{attribute 'qualified_only'}
VAR_GLOBAL
	//Inputs
	DI_E0_0     AT%I*	:BOOL;
	DI_E0_1		AT%I*	:BOOL;
	
	DI_E50_0	AT%I*	:BOOL;
	DI_E50_1	AT%I*	:BOOL;
	DI_E50_2	AT%I*	:BOOL;
	
	DI_E1050_0	AT%I*	:BOOL;
	DI_E1050_1	AT%I*	:BOOL;
	DI_E1050_2	AT%I*	:BOOL;
	DI_E1050_3	AT%I*	:BOOL;
	DI_E1050_4	AT%I*	:BOOL;
	DI_E1050_5	AT%I*	:BOOL;
	
	DI_E1051_0	AT%I*	:BOOL;
	DI_E1051_1	AT%I*	:BOOL;
	DI_E1051_2	AT%I*	:BOOL;
	DI_E1051_3	AT%I*	:BOOL;
	
	DI_E1052_0	AT%I*	:BOOL;
	DI_E1052_1	AT%I*	:BOOL;
	DI_E1052_2	AT%I*	:BOOL;
	DI_E1052_3	AT%I*	:BOOL;
	DI_E1052_4	AT%I*	:BOOL;
	DI_E1052_5	AT%I*	:BOOL;
	DI_E1052_6	AT%I*	:BOOL;
	DI_E1052_7	AT%I*	:BOOL;
	
	
	//Outputs
	DQ_A0_0		AT%Q*	:BOOL;
	DQ_A0_1		AT%Q*	:BOOL;
	
	DQ_A50_0	AT%Q*	:BOOL;
	DQ_A50_1	AT%Q*	:BOOL;
	DQ_A50_2	AT%Q*	:BOOL;
	DQ_A50_3	AT%Q*	:BOOL;
	DQ_A50_4	AT%Q*	:BOOL;
	DQ_A50_5	AT%Q*	:BOOL;
	
	DQ_A1050_0	AT%Q*	:BOOL;
	DQ_A1050_1	AT%Q*	:BOOL;
	DQ_A1050_2	AT%Q*	:BOOL;
	DQ_A1050_3	AT%Q*	:BOOL;
	DQ_A1050_4	AT%Q*	:BOOL;
	DQ_A1050_5	AT%Q*	:BOOL;
	DQ_A1050_6	AT%Q*	:BOOL;
	DQ_A1050_7	AT%Q*	:BOOL;
	
	DQ_A1051_0	AT%Q*	:BOOL;
	DQ_A1051_1	AT%Q*	:BOOL;
	DQ_A1051_2	AT%Q*	:BOOL;
	DQ_A1051_3	AT%Q*	:BOOL;
	DQ_A1051_4	AT%Q*	:BOOL;
	DQ_A1051_5	AT%Q*	:BOOL;
	DQ_A1051_6	AT%Q*	:BOOL;
	DQ_A1051_7	AT%Q*	:BOOL;
	
	
END_VAR

(* stored: Version 1.1.0.1
   GVL GVL_IO: Id {20afe2e4-1740-49e0-8b0a-03a379c1c35b} *)
